Fanuc KAREL source: KO00071.KL

PROGRAM KO00071
%NOLOCKGROUP
%ENVIRONMENT MIR
VAR
  P1: XYZWPREXT
  P2: XYZWPR
  F: BOOLEAN
  OUT: XYZWPREXT
BEGIN
  F = TRUE
  OUT = MIRROR(P1, P2, F)
END KO00071
